(* IEC 61131-3 sources: nautilus/examples/well-site, 3 files *)

(* ---- types.st ---- *)
(* The UDTs a well site is made of. Each site asset is ONE struct tag, so
   the scene binds a whole asset by name (WL101, R101) and reads its
   members. A root .st with no PROGRAM is a library: `type: Well` in the
   manifest resolves against it. *)

TYPE
  Motor : STRUCT
    Run     : BOOL;   (* command *)
    Running : BOOL;   (* feedback *)
    Fault   : BOOL;
    Speed   : REAL;   (* % *)
    Hours   : REAL;
  END_STRUCT;

  (* A production well: the submersible pump, and the water in the casing.
     Depths are metres below grade, so a bigger number is less water. *)
  Well : STRUCT
    Pump   : Motor;
    Depth  : REAL;    (* pumping water level, m below grade *)
    Static : REAL;    (* resting water level, m below grade *)
    Flow   : REAL;    (* at the wellhead, L/s *)
    (* the alarm rules' bits — rules match one level of members, so the
       pump's fault is mirrored here *)
    LL     : BOOL;    (* drawn down past the limit *)
    Fault  : BOOL;    (* = Pump.Fault *)
  END_STRUCT;

  Meter : STRUCT
    Flow  : REAL;     (* L/s *)
    Total : REAL;     (* m3 *)
  END_STRUCT;

  Valve : STRUCT
    Cmd   : REAL;     (* % open command *)
    Pos   : REAL;     (* % open feedback *)
    Fault : BOOL;     (* position disagrees with command *)
  END_STRUCT;

  Tank : STRUCT
    Level : REAL;     (* % *)
    TempC : REAL;
    HH    : BOOL;
    LL    : BOOL;
  END_STRUCT;

  (* Hypochlorite feed: a day tank and a dosing pump, as a UDT of UDTs,
     so the scene places the skid as one node and its parts read
     CL101.Tank and CL101.Pump (docs/design/spatial-hmi.md §3d). *)
  ChemFeed : STRUCT
    Tank     : Tank;
    Pump     : Motor;
    Residual : REAL;  (* mg/L free chlorine at the injection point *)
    Low      : BOOL;  (* residual under the limit *)
    Fault    : BOOL;  (* = Pump.Fault *)
  END_STRUCT;
END_TYPE

(* ---- control.st ---- *)
PROGRAM Control
(* The site's control logic: the well pump fills the reservoir between
   two levels, the discharge valve opens with the pump, the hypochlorite
   pump doses while water moves, and the limit bits the alarms claim. *)
VAR_EXTERNAL
    WL101 : Well;
    FIT101 : Meter;
    FCV101 : Valve;
    CL101 : ChemFeed;
    R101 : Tank;
    StartLevel : REAL;
    StopLevel : REAL;
    MaxDepth : REAL;
    ResidualLow : REAL;
    ControlDtS : REAL;
END_VAR
VAR
    valveDisagreeS : REAL;   (* how long the valve has been off its command *)
END_VAR

(* the drawdown limit, with hysteresis so the alarm holds while the well
   recovers instead of chattering on the limit *)
IF WL101.Depth > MaxDepth THEN
    WL101.LL := TRUE;
ELSIF WL101.Depth < MaxDepth - 0.3 THEN
    WL101.LL := FALSE;
END_IF;
WL101.Fault := WL101.Pump.Fault;
CL101.Fault := CL101.Pump.Fault;

(* well pump seal-in on reservoir level; never on a fault, never when the
   water has been drawn down past the limit *)
IF WL101.Pump.Fault OR WL101.LL THEN
    WL101.Pump.Run := FALSE;
ELSIF R101.Level < StartLevel THEN
    WL101.Pump.Run := TRUE;
ELSIF R101.Level > StopLevel THEN
    WL101.Pump.Run := FALSE;
END_IF;
IF WL101.Pump.Running THEN
    WL101.Pump.Hours := WL101.Pump.Hours + ControlDtS / 3600.0;
END_IF;

(* the discharge valve opens with the pump's run command; a valve that is
   still off its command after a full stroke's worth of time is stuck *)
IF WL101.Pump.Run THEN
    FCV101.Cmd := 100.0;
ELSE
    FCV101.Cmd := 0.0;
END_IF;
IF ABS(FCV101.Cmd - FCV101.Pos) > 10.0 THEN
    valveDisagreeS := valveDisagreeS + ControlDtS;
ELSE
    valveDisagreeS := 0.0;
END_IF;
FCV101.Fault := valveDisagreeS > 8.0;

(* dose while the meter sees flow *)
CL101.Pump.Run := FIT101.Flow > 0.5 AND NOT CL101.Pump.Fault AND CL101.Tank.Level > 2.0;
CL101.Low := FIT101.Flow > 0.5 AND CL101.Residual < ResidualLow;
CL101.Tank.LL := CL101.Tank.Level < 10.0;

R101.HH := R101.Level > 95.0;
R101.LL := R101.Level < 10.0;
END_PROGRAM

(* ---- sim.st ---- *)
PROGRAM Sim
(* Stands in for the field: the aquifer, the pipe, the reservoir and the
   chlorine, plus switches to make something go wrong on demand. *)
VAR_EXTERNAL
    WL101 : Well;
    FIT101 : Meter;
    FCV101 : Valve;
    CL101 : ChemFeed;
    R101 : Tank;
    SimDtS : REAL;
    InjectPumpFault : BOOL;
    InjectDrought : BOOL;
END_VAR
VAR CONSTANT
    WellMaxLps : REAL := 12.0;     (* at 100 % speed *)
    DrawdownMPerLps : REAL := 0.06; (* the cone of depression, per L/s *)
    AquiferTauS : REAL := 20.0;    (* how fast the level follows the pumping *)
    ReservoirM3 : REAL := 6.0;     (* tiny, so a fill is minutes, not hours *)
    TownLps : REAL := 5.0;         (* what the town draws, steadily *)
    ValveRatePctS : REAL := 20.0;
    PumpRampPctS : REAL := 25.0;
    DayTankPctPerS : REAL := 0.02;
END_VAR
VAR
    target : REAL;
    step : REAL;
END_VAR

(* the well pump *)
WL101.Pump.Fault := InjectPumpFault;
WL101.Pump.Running := WL101.Pump.Run AND NOT WL101.Pump.Fault;
IF WL101.Pump.Running THEN
    WL101.Pump.Speed := MIN(WL101.Pump.Speed + PumpRampPctS * SimDtS, 100.0);
ELSE
    WL101.Pump.Speed := MAX(WL101.Pump.Speed - PumpRampPctS * SimDtS, 0.0);
END_IF;
WL101.Flow := WL101.Pump.Speed / 100.0 * WellMaxLps;

(* the aquifer: the water level settles toward static plus the drawdown
   the flow earns, with a lag; a drought sinks the static level *)
IF InjectDrought THEN
    WL101.Static := 1.15;
ELSE
    WL101.Static := 0.45;
END_IF;
target := WL101.Static + DrawdownMPerLps * WL101.Flow;
WL101.Depth := WL101.Depth + (target - WL101.Depth) * SimDtS / AquiferTauS;

(* the discharge valve strokes toward its command *)
step := ValveRatePctS * SimDtS;
FCV101.Pos := FCV101.Pos + LIMIT(-step, FCV101.Cmd - FCV101.Pos, step);

(* the meter sees what the valve passes *)
FIT101.Flow := WL101.Flow * FCV101.Pos / 100.0;
FIT101.Total := FIT101.Total + FIT101.Flow * SimDtS / 1000.0;

(* the reservoir: fills from the well, drains to the town *)
R101.Level := LIMIT(0.0, R101.Level + (FIT101.Flow - TownLps) * SimDtS / ReservoirM3 / 10.0, 100.0);
R101.TempC := 14.0;

(* hypochlorite: the dosing pump draws the day tank down and holds the
   residual while it runs; the residual decays when it stops *)
CL101.Pump.Running := CL101.Pump.Run AND NOT CL101.Pump.Fault;
IF CL101.Pump.Running THEN
    CL101.Pump.Speed := 100.0;
    CL101.Tank.Level := MAX(CL101.Tank.Level - DayTankPctPerS * SimDtS, 0.0);
    CL101.Residual := CL101.Residual + (1.2 - CL101.Residual) * SimDtS / 15.0;
ELSE
    CL101.Pump.Speed := 0.0;
    CL101.Residual := MAX(CL101.Residual - 0.05 * SimDtS, 0.0);
END_IF;
END_PROGRAM
